PROGRAM PRG_TEST
VAR
    fb_PPEPS_Tests : FB_PPEPS_Tests;
    {attribute 'TcNcAxis' := '
        .fbAxisRef[1] := Axis_HomeToCenter_Test1;
        .fbAxisRef[2] := Axis_HomeToCenter_Test2;
        .fbAxisRef[3] := Axis_HomeToCenter_Test3;
        .fbAxisRef[4] := Axis_HomeToCenter_Test4;
        .fbAxisRef[5] := Axis_HomeToCenter_Test5;
    '}
    fb_HomeToCenter_Tests : FB_HomeToCenter_Tests;
END_VAR

TcUnit.Run();

END_PROGRAM

(* stored: Version 1.1.0.1
   POU PRG_TEST: Id {8dc7f58a-f85f-4fee-87b3-7c48ea7c69af}, SpecialFunc None *)
